Universal Robots URScript: letra_G.script

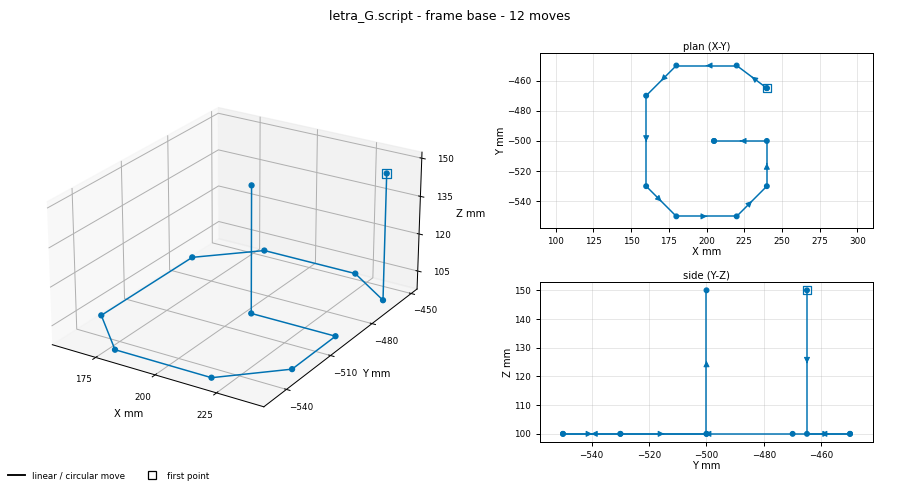
[picture p0: tool path of letra_G.script in frame base, 12 of 12 moves have a stored position in this frame; points joined in program order, loops and branches not executed]
# Letra G - Garcia
movel(p[0.240, -0.465, 0.150, 3.1416, 0, 0], a=0.5, v=0.1)
movel(p[0.240, -0.465, 0.100, 3.1416, 0, 0], a=0.5, v=0.1)
movel(p[0.220, -0.450, 0.100, 3.1416, 0, 0], a=0.5, v=0.1)
movel(p[0.180, -0.450, 0.100, 3.1416, 0, 0], a=0.5, v=0.1)
movel(p[0.160, -0.470, 0.100, 3.1416, 0, 0], a=0.5, v=0.1)
movel(p[0.160, -0.530, 0.100, 3.1416, 0, 0], a=0.5, v=0.1)
movel(p[0.180, -0.550, 0.100, 3.1416, 0, 0], a=0.5, v=0.1)
movel(p[0.220, -0.550, 0.100, 3.1416, 0, 0], a=0.5, v=0.1)
movel(p[0.240, -0.530, 0.100, 3.1416, 0, 0], a=0.5, v=0.1)
movel(p[0.240, -0.500, 0.100, 3.1416, 0, 0], a=0.5, v=0.1)
movel(p[0.205, -0.500, 0.100, 3.1416, 0, 0], a=0.5, v=0.1)
movel(p[0.205, -0.500, 0.150, 3.1416, 0, 0], a=0.5, v=0.1)
